(* IEC 61131-3 sources: axsharp/src/AXSharp.compiler/tests/AXSharp.Compiler.CsTests/samples/sourcefile/src/sub, 1 file *)

(* ---- widget.st ---- *)
CLASS widget

END_CLASS

TYPE
    Gadget : STRUCT
        running : BOOL;
    END_STRUCT;
END_TYPE

TYPE
    Shade : (Light, Dark) := Light;
END_TYPE

INTERFACE PUBLIC IWidget

END_INTERFACE
